FUNCTION_BLOCK ArmReset (* Basic Function Block Type *)
  (* Standard: 61499-2 *)
  (* Version 0.0, 7/2/2026, Template *)
  PACKAGE Main;
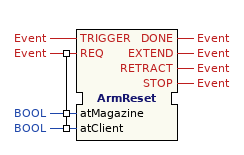
  EVENT_INPUT
    TRIGGER;
    REQ WITH atMagazine, atClient; (* Normal Execution Request *)
  END_EVENT
  EVENT_OUTPUT
    DONE;
    EXTEND;
    RETRACT;
    STOP;
  END_EVENT
  VAR_INPUT
    atMagazine : BOOL; (* Input event qualifier *)
    atClient : BOOL;
  END_VAR
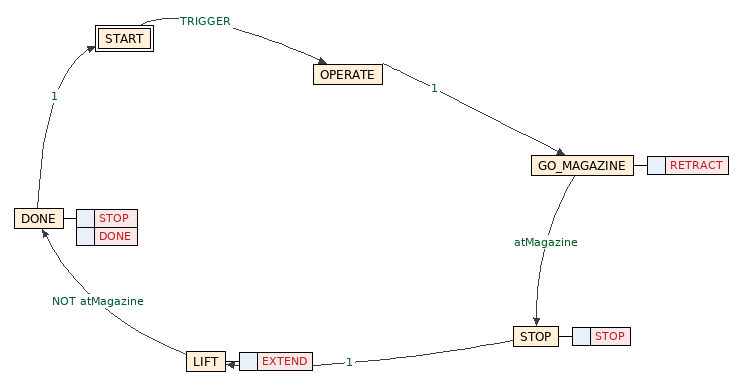
  EC_STATES
    START; (* Initial State *)
    OPERATE;
    GO_MAGAZINE : -> RETRACT;
    STOP : -> STOP;
    LIFT : -> EXTEND;
    DONE : -> STOP, -> DONE;
  END_STATES
  EC_TRANSITIONS
    START TO OPERATE := TRIGGER;
    OPERATE TO GO_MAGAZINE := 1;
    GO_MAGAZINE TO STOP := atMagazine;
    STOP TO LIFT := 1;
    LIFT TO DONE := NOT atMagazine;
    DONE TO START := 1;
  END_TRANSITIONS
  ALGORITHM INIT IN ST: (* Initialization algorithm *)
;
  END_ALGORITHM
  ALGORITHM REQ IN ST: (* Normally executed algorithm *)
;
  END_ALGORITHM
END_FUNCTION_BLOCK
